Fanuc KAREL source: KD00020.KL

PROGRAM KD00020
%NOLOCKGROUP
VAR
  I: INTEGER
  J: INTEGER
  B: BOOLEAN
  R: REAL
  S: STRING[80]
BEGIN
  GO TO done
done:: I = 1
END KD00020
